{attribute 'linkalways'}
{attribute 'no_explicit_call' := 'Use the methods of this class'}
{attribute 'enable_dynamic_creation'}
FUNCTION_BLOCK SimulatorLink
VAR
	cycle : UDINT;
	lastSequence : UDINT;
	silentCycles : UDINT;
	_isConnected : BOOL;
END_VAR

METHOD Execute
cycle := cycle + 1;
SimulatorIo.command.version := Constants.SIMULATOR_PROTOCOL_VERSION;
SimulatorIo.command.cycle := cycle;
SimulatorIo.command.plcTimeInNs := F_GetSystemTime() * 100;

IF SimulatorIo.feedback.sequence <> lastSequence THEN
	lastSequence := SimulatorIo.feedback.sequence;
	silentCycles := 0;
ELSIF silentCycles < Constants.SIMULATOR_TIMEOUT_IN_CYCLES THEN
	silentCycles := silentCycles + 1;
END_IF

_isConnected := SimulatorIo.feedback.version = Constants.SIMULATOR_PROTOCOL_VERSION
	AND silentCycles < Constants.SIMULATOR_TIMEOUT_IN_CYCLES;
END_METHOD

PROPERTY IsConnected : BOOL
GET
IsConnected := _isConnected;
END_GET
END_PROPERTY

END_FUNCTION_BLOCK

(* stored: Version 1.1.0.1, ProductVersion 3.1.4026.12
   POU SimulatorLink: Id {a462f8c5-672d-5d13-8abd-5a10e743d669}, SpecialFunc None
   Method Execute: Id {6720d030-624d-54b3-ab2f-48c7aca86e3c}
   Property IsConnected: Id {14dc0167-7af7-5b4f-bb02-e46a92a05599}
   Get Get: Id {afc8f24c-0732-53bc-a83c-5208f1ad3ce1} *)
